// TwinCAT 3 PLC project ExperimentSequencerTests
// ProgramVersion: 3.1.4026.22
// libraries:
//   Tc2_Standard, * (Beckhoff Automation GmbH)
//   Tc2_System, * (Beckhoff Automation GmbH)
// project tree:
//   ExperimentSequencer/DUTs/ E_SeqState.TcDUT
//   ExperimentSequencer/tests/GVLs/ GVL_SEQ.TcGVL
//   ExperimentSequencer/POUs/ FB_ExperimentSequencerCore.TcPOU, PRG_ExperimentSequencer.TcPOU
//   ExperimentSequencer/tests/POUs/ PRG_ExperimentSequencerTests.TcPOU
//   ExperimentSequencer/tests/ TestTask.TcTTO
// real-time tasks:
//   TASK DriveStateTestTask: cycle T#10ms, priority 1, ADS port 350
//   TASK TestTask: cycle T#10ms, priority 2, ADS port 351

CONFIGURATION ExperimentSequencerTests
    RESOURCE PLC ON TwinCAT3
        TASK TestTask(INTERVAL := T#10ms, PRIORITY := 2);
        PROGRAM PRG_ExperimentSequencer WITH TestTask : PRG_ExperimentSequencer;
        PROGRAM PRG_ExperimentSequencerTests WITH TestTask : PRG_ExperimentSequencerTests;
    END_RESOURCE
END_CONFIGURATION

// ---- ExperimentSequencer/DUTs/E_SeqState.TcDUT
{attribute 'qualified_only'}
{attribute 'strict'}
TYPE E_SeqState :
(
    IDLE := 0,          (* Waiting. Outputs zeroed. *)
    PLAYING := 10,      (* Table playback active. *)
    COMPLETE := 20,     (* Playback complete, outputs held until rearm. *)
    FAULT := 90         (* Invalid input detected, reset edge required. *)
);
END_TYPE

// ---- ExperimentSequencer/tests/GVLs/GVL_SEQ.TcGVL
{attribute 'qualified_only'}
VAR_GLOBAL CONSTANT
    N_REF_MAX : UDINT := 8;
    N_FF_MAX : UDINT := 8;
    N_DIST_MAX : UDINT := 8;
END_VAR

VAR_GLOBAL
    refValue : LREAL := 0.0;
    ffValue : LREAL := 0.0;
    distValue : LREAL := 0.0;
    refTable : ARRAY[0..N_REF_MAX - 1] OF LREAL;
    ffTable : ARRAY[0..N_FF_MAX - 1] OF LREAL;
    distTable : ARRAY[0..N_DIST_MAX - 1] OF LREAL;
    tableLen : UDINT := 0;
    idx : UDINT := 0;
    repeatCount : UDINT := 1;
    trialIndex : UDINT := 0;
    resetReq : BOOL := FALSE;
    experimentActive : BOOL := FALSE;
    playbackDone : BOOL := FALSE;
    seqError : BOOL := FALSE;
    seqState : E_SeqState := E_SeqState.IDLE;
    tableLenClamped : UDINT := 0;
END_VAR

// ---- ExperimentSequencer/POUs/PRG_ExperimentSequencer.TcPOU
PROGRAM PRG_ExperimentSequencer
VAR
    tableIdxDint : DINT := 0;
    tableLenLocal : UDINT := 0;
    tableLenMaxLocal : UDINT := 0;
    refSample : LREAL := 0.0;
    ffSample : LREAL := 0.0;
    distSample : LREAL := 0.0;
    fbSequencerCore : FB_ExperimentSequencerCore;
END_VAR

tableLenMaxLocal := GVL_SEQ.N_REF_MAX;
IF GVL_SEQ.N_FF_MAX < tableLenMaxLocal THEN
    tableLenMaxLocal := GVL_SEQ.N_FF_MAX;
END_IF
IF GVL_SEQ.N_DIST_MAX < tableLenMaxLocal THEN
    tableLenMaxLocal := GVL_SEQ.N_DIST_MAX;
END_IF

tableLenLocal := GVL_SEQ.tableLen;
IF tableLenLocal > tableLenMaxLocal THEN
    tableLenLocal := tableLenMaxLocal;
END_IF
GVL_SEQ.tableLenClamped := tableLenLocal;

refSample := 0.0;
ffSample := 0.0;
distSample := 0.0;
IF fbSequencerCore.idx < tableLenLocal THEN
    tableIdxDint := UDINT_TO_DINT(fbSequencerCore.idx);
    refSample := GVL_SEQ.refTable[tableIdxDint];
    ffSample := GVL_SEQ.ffTable[tableIdxDint];
    distSample := GVL_SEQ.distTable[tableIdxDint];
END_IF

fbSequencerCore(
    resetRequest := GVL_SEQ.resetReq,
    experimentActive := GVL_SEQ.experimentActive,
    tableLen := tableLenLocal,
    repeatCount := GVL_SEQ.repeatCount,
    refSample := refSample,
    ffSample := ffSample,
    distSample := distSample
);

GVL_SEQ.refValue := fbSequencerCore.refValue;
GVL_SEQ.ffValue := fbSequencerCore.ffValue;
GVL_SEQ.distValue := fbSequencerCore.distValue;
GVL_SEQ.playbackDone := fbSequencerCore.playbackDone;
GVL_SEQ.seqError := fbSequencerCore.seqError;
GVL_SEQ.seqState := fbSequencerCore.seqState;
GVL_SEQ.idx := fbSequencerCore.idx;
GVL_SEQ.trialIndex := fbSequencerCore.trialIndex;

END_PROGRAM

// ---- ExperimentSequencer/POUs/FB_ExperimentSequencerCore.TcPOU
FUNCTION_BLOCK FB_ExperimentSequencerCore
VAR_INPUT
    resetRequest : BOOL;
    experimentActive : BOOL;
    tableLen : UDINT;
    repeatCount : UDINT;
    refSample : LREAL;
    ffSample : LREAL;
    distSample : LREAL;
END_VAR
VAR_OUTPUT
    refValue : LREAL := 0.0;
    ffValue : LREAL := 0.0;
    distValue : LREAL := 0.0;
    playbackDone : BOOL := FALSE;
    seqError : BOOL := FALSE;
    seqState : E_SeqState := E_SeqState.IDLE;
    idx : UDINT := 0;
    trialIndex : UDINT := 0;
END_VAR
VAR
    experimentActivePrev : BOOL := FALSE;
    resetRequestPrev : BOOL := FALSE;
    resetEdge : BOOL := FALSE;
    startEdge : BOOL := FALSE;
    zeroOutputsThisScan : BOOL := FALSE;
    resetProgressThisScan : BOOL := FALSE;
END_VAR

zeroOutputsThisScan := FALSE;
resetProgressThisScan := FALSE;
resetEdge := resetRequest AND NOT resetRequestPrev;
startEdge := experimentActive AND NOT experimentActivePrev;

IF resetEdge THEN
    resetProgressThisScan := TRUE;
    zeroOutputsThisScan := TRUE;
    seqState := E_SeqState.IDLE;

ELSE
    CASE seqState OF
        E_SeqState.IDLE:
            zeroOutputsThisScan := TRUE;

            IF startEdge THEN
                IF (tableLen = 0) OR (repeatCount = 0) THEN
                    seqState := E_SeqState.FAULT;
                ELSE
                    resetProgressThisScan := TRUE;
                    seqState := E_SeqState.PLAYING;
                END_IF
            END_IF

        E_SeqState.PLAYING:
            IF NOT experimentActive THEN
                resetProgressThisScan := TRUE;
                zeroOutputsThisScan := TRUE;
                seqState := E_SeqState.IDLE;
            ELSIF idx < tableLen THEN
                refValue := refSample;
                ffValue := ffSample;
                distValue := distSample;
                idx := idx + 1;

                IF idx >= tableLen THEN
                    IF trialIndex >= (repeatCount - 1) THEN
                        playbackDone := TRUE;
                        seqState := E_SeqState.COMPLETE;
                    ELSE
                        idx := 0;
                        trialIndex := trialIndex + 1;
                    END_IF
                END_IF
            END_IF

        E_SeqState.COMPLETE:
            IF NOT experimentActive THEN
                resetProgressThisScan := TRUE;
                zeroOutputsThisScan := TRUE;
                seqState := E_SeqState.IDLE;
            END_IF

        E_SeqState.FAULT:
            resetProgressThisScan := TRUE;
            zeroOutputsThisScan := TRUE;
    END_CASE
END_IF

IF resetProgressThisScan THEN
    idx := 0;
    trialIndex := 0;
END_IF
IF zeroOutputsThisScan THEN
    refValue := 0.0;
    ffValue := 0.0;
    distValue := 0.0;
    playbackDone := FALSE;
END_IF

seqError := (seqState = E_SeqState.FAULT);
experimentActivePrev := experimentActive;
resetRequestPrev := resetRequest;

END_FUNCTION_BLOCK

// ---- ExperimentSequencer/tests/POUs/PRG_ExperimentSequencerTests.TcPOU
PROGRAM PRG_ExperimentSequencerTests
VAR
    stage : UINT := 0;
    testsExecuted : BOOL := FALSE;
    testsPassed : BOOL := FALSE;
    failureCount : UDINT := 0;
END_VAR

IF NOT testsExecuted THEN
    CASE stage OF
        0:
            GVL_SEQ.tableLen := 9;
            GVL_SEQ.repeatCount := 1;
            GVL_SEQ.experimentActive := FALSE;
            GVL_SEQ.resetReq := FALSE;
            stage := 1;

        1:
            IF (GVL_SEQ.tableLenClamped <> 8) OR (GVL_SEQ.seqState <> E_SeqState.IDLE) THEN
                failureCount := failureCount + 1;
            END_IF
            GVL_SEQ.refTable[0] := 1.0;
            GVL_SEQ.refTable[1] := 2.0;
            GVL_SEQ.refTable[2] := 3.0;
            GVL_SEQ.ffTable[0] := 10.0;
            GVL_SEQ.ffTable[1] := 20.0;
            GVL_SEQ.ffTable[2] := 30.0;
            GVL_SEQ.distTable[0] := 100.0;
            GVL_SEQ.distTable[1] := 200.0;
            GVL_SEQ.distTable[2] := 300.0;
            GVL_SEQ.tableLen := 3;
            GVL_SEQ.repeatCount := 2;
            GVL_SEQ.experimentActive := TRUE;
            stage := 2;

        2:
            IF (GVL_SEQ.seqState <> E_SeqState.PLAYING)
                OR (GVL_SEQ.idx <> 0) OR (GVL_SEQ.trialIndex <> 0)
                OR GVL_SEQ.playbackDone OR (GVL_SEQ.refValue <> 0.0) THEN
                failureCount := failureCount + 1;
            END_IF
            stage := 3;

        3:
            IF (GVL_SEQ.idx <> 1) OR (GVL_SEQ.trialIndex <> 0)
                OR (GVL_SEQ.refValue <> 1.0) OR (GVL_SEQ.ffValue <> 10.0)
                OR (GVL_SEQ.distValue <> 100.0) OR GVL_SEQ.playbackDone THEN
                failureCount := failureCount + 1;
            END_IF
            stage := 4;

        4:
            IF (GVL_SEQ.idx <> 2) OR (GVL_SEQ.refValue <> 2.0)
                OR (GVL_SEQ.ffValue <> 20.0) OR (GVL_SEQ.distValue <> 200.0) THEN
                failureCount := failureCount + 1;
            END_IF
            stage := 5;

        5:
            IF (GVL_SEQ.idx <> 0) OR (GVL_SEQ.trialIndex <> 1)
                OR (GVL_SEQ.refValue <> 3.0) OR GVL_SEQ.playbackDone THEN
                failureCount := failureCount + 1;
            END_IF
            stage := 6;

        6:
            IF (GVL_SEQ.idx <> 1) OR (GVL_SEQ.trialIndex <> 1)
                OR (GVL_SEQ.refValue <> 1.0) THEN
                failureCount := failureCount + 1;
            END_IF
            stage := 7;

        7:
            IF (GVL_SEQ.idx <> 2) OR (GVL_SEQ.refValue <> 2.0) THEN
                failureCount := failureCount + 1;
            END_IF
            stage := 8;

        8:
            IF (GVL_SEQ.seqState <> E_SeqState.COMPLETE)
                OR (GVL_SEQ.idx <> 3) OR (GVL_SEQ.trialIndex <> 1)
                OR NOT GVL_SEQ.playbackDone OR (GVL_SEQ.refValue <> 3.0) THEN
                failureCount := failureCount + 1;
            END_IF
            GVL_SEQ.experimentActive := FALSE;
            stage := 9;

        9:
            IF (GVL_SEQ.seqState <> E_SeqState.IDLE)
                OR (GVL_SEQ.idx <> 0) OR (GVL_SEQ.trialIndex <> 0)
                OR GVL_SEQ.playbackDone OR (GVL_SEQ.refValue <> 0.0)
                OR (GVL_SEQ.ffValue <> 0.0) OR (GVL_SEQ.distValue <> 0.0) THEN
                failureCount := failureCount + 1;
            END_IF
            GVL_SEQ.tableLen := 3;
            GVL_SEQ.repeatCount := 1;
            GVL_SEQ.experimentActive := TRUE;
            stage := 10;

        10:
            IF (GVL_SEQ.seqState <> E_SeqState.PLAYING) OR (GVL_SEQ.idx <> 0) THEN
                failureCount := failureCount + 1;
            END_IF
            stage := 11;

        11:
            IF (GVL_SEQ.idx <> 1) OR (GVL_SEQ.refValue <> 1.0) THEN
                failureCount := failureCount + 1;
            END_IF
            GVL_SEQ.experimentActive := FALSE;
            stage := 12;

        12:
            IF (GVL_SEQ.seqState <> E_SeqState.IDLE)
                OR (GVL_SEQ.idx <> 0) OR (GVL_SEQ.trialIndex <> 0)
                OR GVL_SEQ.playbackDone OR (GVL_SEQ.refValue <> 0.0) THEN
                failureCount := failureCount + 1;
            END_IF
            GVL_SEQ.tableLen := 0;
            GVL_SEQ.repeatCount := 1;
            GVL_SEQ.experimentActive := TRUE;
            stage := 13;

        13:
            IF (GVL_SEQ.seqState <> E_SeqState.FAULT) OR NOT GVL_SEQ.seqError
                OR GVL_SEQ.playbackDone OR (GVL_SEQ.refValue <> 0.0) THEN
                failureCount := failureCount + 1;
            END_IF
            GVL_SEQ.resetReq := TRUE;
            stage := 14;

        14:
            IF (GVL_SEQ.seqState <> E_SeqState.IDLE) OR GVL_SEQ.seqError
                OR (GVL_SEQ.idx <> 0) OR (GVL_SEQ.trialIndex <> 0) THEN
                failureCount := failureCount + 1;
            END_IF
            GVL_SEQ.resetReq := FALSE;
            GVL_SEQ.experimentActive := FALSE;
            stage := 15;

        15:
            GVL_SEQ.resetReq := TRUE;
            GVL_SEQ.experimentActive := TRUE;
            stage := 16;

        16:
            IF (GVL_SEQ.seqState <> E_SeqState.IDLE) OR GVL_SEQ.seqError
                OR (GVL_SEQ.idx <> 0) OR (GVL_SEQ.trialIndex <> 0)
                OR GVL_SEQ.playbackDone THEN
                failureCount := failureCount + 1;
            END_IF
            GVL_SEQ.resetReq := FALSE;
            GVL_SEQ.experimentActive := FALSE;
            stage := 17;

        17:
            GVL_SEQ.tableLen := 3;
            GVL_SEQ.repeatCount := 0;
            GVL_SEQ.experimentActive := TRUE;
            stage := 18;

        18:
            IF (GVL_SEQ.seqState <> E_SeqState.FAULT) OR NOT GVL_SEQ.seqError
                OR (GVL_SEQ.idx <> 0) OR (GVL_SEQ.trialIndex <> 0)
                OR GVL_SEQ.playbackDone OR (GVL_SEQ.refValue <> 0.0) THEN
                failureCount := failureCount + 1;
            END_IF
            GVL_SEQ.resetReq := TRUE;
            stage := 19;

        19:
            IF (GVL_SEQ.seqState <> E_SeqState.IDLE) OR GVL_SEQ.seqError
                OR (GVL_SEQ.idx <> 0) OR (GVL_SEQ.trialIndex <> 0)
                OR GVL_SEQ.playbackDone THEN
                failureCount := failureCount + 1;
            END_IF
            GVL_SEQ.resetReq := FALSE;
            GVL_SEQ.experimentActive := FALSE;
            testsExecuted := TRUE;
            testsPassed := (failureCount = 0);
    END_CASE
END_IF

END_PROGRAM
